(* IEC 61131-3 sources: trust-platform/conformance/cases/enums/cfm_enums_variant_assignment_001, 1 file *)

(* ---- program.st ---- *)
TYPE Phase :
(
    IDLE := 0,
    RUNNING := 1,
    DONE := 2
);
END_TYPE

PROGRAM Main
VAR
    state : Phase := Phase#IDLE;
    is_running : BOOL := FALSE;
END_VAR

state := RUNNING;
is_running := state = RUNNING;
END_PROGRAM
